Fanuc KAREL source: KA00114.KL

PROGRAM KA00114
%NOLOCKGROUP
VAR
  SRC: CONFIG
  DST: XYZWPR
BEGIN
  SRC.CFG_FLIP = TRUE
  DST = SRC
END KA00114
